Fanuc KAREL source: kb00104.KL

-- PROVISIONAL review KL for V940-1; original PC SHA256 8b68e5b2633bbdf2579a3230d504adc9b67411bf5a92f7e3906b6d5856ea7c3f
-- Incomplete behavior may be omitted. Consult companion uncertainty JSON. Do not deploy.
PROGRAM KB00104
%NOLOCKGROUP
BEGIN
  -- V9_ZERO_TABLE_METADATA_HINT layout=0002_ascii; no indexed target words; source/name/runtime held
  -- UNRESOLVED_PC offsets 5-16; opcodes 2E,23
  -- UNRESOLVED_PC offsets 21-30; opcodes 3F,75
  -- UNRESOLVED_PC offsets 35-42; opcodes 9D,23
  -- UNRESOLVED_PC offsets 47-54; opcodes 9D,23
  -- UNRESOLVED_PC offsets 59-66; opcodes 9D,23
  -- UNRESOLVED_PC offsets 71-78; opcodes 9D,23
  -- UNRESOLVED_PC offsets 83-90; opcodes 9D,23
  -- UNRESOLVED_PC offsets 95-102; opcodes 9D,23
  -- UNRESOLVED_PC offsets 107-114; opcodes 9D,23
  -- UNRESOLVED_PC offsets 119-128; opcodes 3F,75
  -- UNRESOLVED_PC offsets 133-140; opcodes 9D,23
  -- UNRESOLVED_PC offsets 145-219; opcodes 27,22,22,2A,22,22,22,22,22,22,22,22,2A,22,31
  -- UNRESOLVED_PC offsets 224-228; opcodes 7F
END KB00104
